{attribute 'reflection'}
FUNCTION_BLOCK FB_Error
VAR_OUTPUT
	bError:		BOOL;
	nErrorID:	UDINT;
	eErrorID:	E_ErrorIDs;
	eErrorSrc:	E_ErrorSrcs;
	sErrorMsg:	STRING(128);
	nState:		INT; //State in dem der Error aufgetreten ist
	
	//{attribute 'instance-path'}
	//{attribute 'no_init'}
	//sSource:	STRING;
END_VAR

METHOD M_Reset
VAR_INPUT
END_VAR
IF bError THEN
	HMI.fbErrorCollector.M_QuitError(eErrorID, eErrorSrc);
	MEMSET(ADR(THIS^), 0, SIZEOF(THIS^));
END_IF
END_METHOD

METHOD M_Set
VAR_INPUT
	nID:	UDINT;
	sMsg:	STRING;
	nState:	INT; //State in dem der Error aufgetreten ist
	eID:	E_ErrorIDs;
	eSrc:	E_ErrorSrcs;
END_VAR
VAR_INST
	
END_VAR
IF NOT bError THEN
	bError := TRUE;
	nErrorID := nID;
	sErrorMsg := sMsg;
	THIS^.nState := nState;
	eErrorID := eID;
	eErrorSrc := eSrc;
	HMI.fbErrorCollector.M_NewError(eID, eSrc, sMsg);
END_IF
END_METHOD

END_FUNCTION_BLOCK

(* stored: Version 1.1.0.1, ProductVersion 3.1.4024.12
   POU FB_Error: Id {643ec9f9-d7f1-4f20-8f55-a071f44f9ecb}, SpecialFunc None
   Method M_Reset: Id {bc054357-f4aa-4638-99d3-83b7f76f5261}
   Method M_Set: Id {6fe6d8ed-fd27-46f4-aaf3-4a28d22d6000} *)
